Fanuc KAREL source: KB00169.KL

PROGRAM KB00169
%NOLOCKGROUP
VAR
  P1: JOINTPOS
  P2: REAL
  P3: INTEGER
BEGIN
  P2 = 1.0
  P3 = 1
  SET_PERCH(P1, P2, P3)
END KB00169
